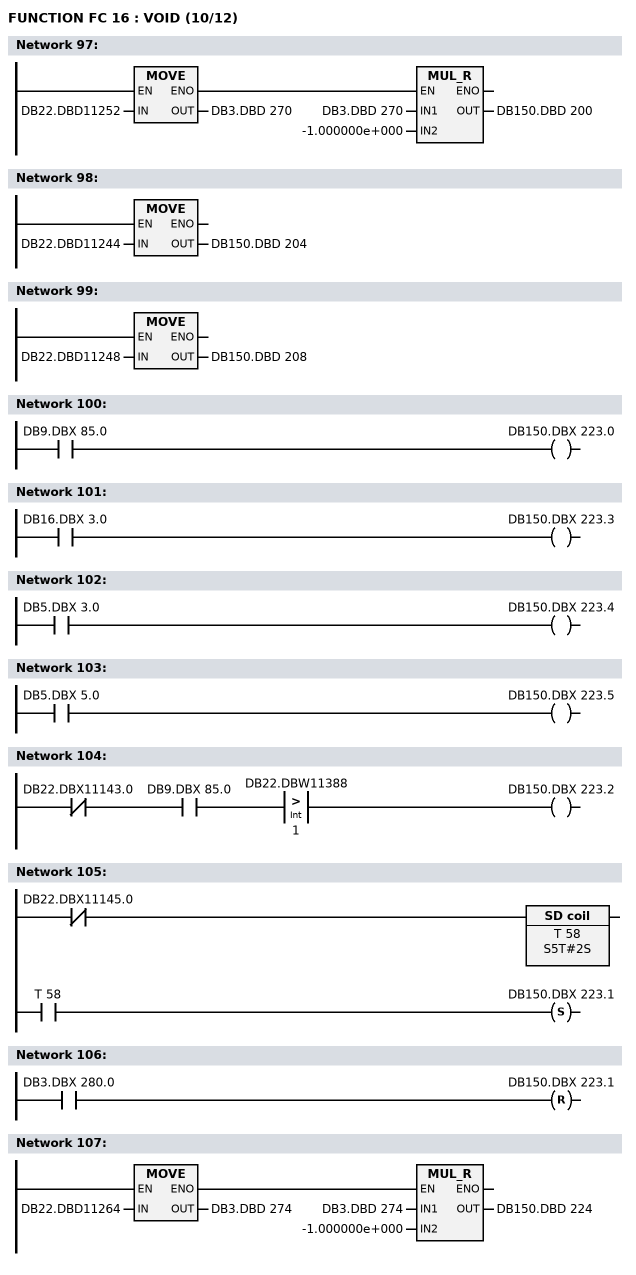

      A(    ;
      L     DB22.DBD11252;
      T     DB3.DBD  270;
      SET   ;
      SAVE  ;
      CLR   ;
      A     BR;
      )     ;
      JNB   M017;
      L     DB3.DBD  270;
      L     -1.000000e+000;
      *R    ;
      T     DB150.DBD  200;
M017: NOP   0;
NETWORK
TITLE =

      L     DB22.DBD11244;
      T     DB150.DBD  204;
      NOP   0;
NETWORK
TITLE =

      L     DB22.DBD11248;
      T     DB150.DBD  208;
      NOP   0;
NETWORK
TITLE =

      A     DB9.DBX   85.0;
      =     DB150.DBX  223.0;
NETWORK
TITLE =

      A     DB16.DBX    3.0;
      =     DB150.DBX  223.3;
NETWORK
TITLE =

      A     DB5.DBX    3.0;
      =     DB150.DBX  223.4;
NETWORK
TITLE =

      A     DB5.DBX    5.0;
      =     DB150.DBX  223.5;
NETWORK
TITLE =

      AN    DB22.DBX11143.0;
      A     DB9.DBX   85.0;
      A(    ;
      L     DB22.DBW11388;
      L     1;
      >I    ;
      )     ;
      =     DB150.DBX  223.2;
NETWORK
TITLE =

      AN    DB22.DBX11145.0;
      L     S5T#2S;
      SD    T     58;
      NOP   0;
      NOP   0;
      NOP   0;
      A     T     58;
      S     DB150.DBX  223.1;
NETWORK
TITLE =

      A     DB3.DBX  280.0;
      R     DB150.DBX  223.1;
NETWORK
TITLE =

      A(    ;
      L     DB22.DBD11264;
      T     DB3.DBD  274;
      SET   ;
      SAVE  ;
      CLR   ;
      A     BR;
      )     ;
      JNB   M018;
      L     DB3.DBD  274;
      L     -1.000000e+000;
      *R    ;
      T     DB150.DBD  224;
M018: NOP   0;
NETWORK
TITLE =
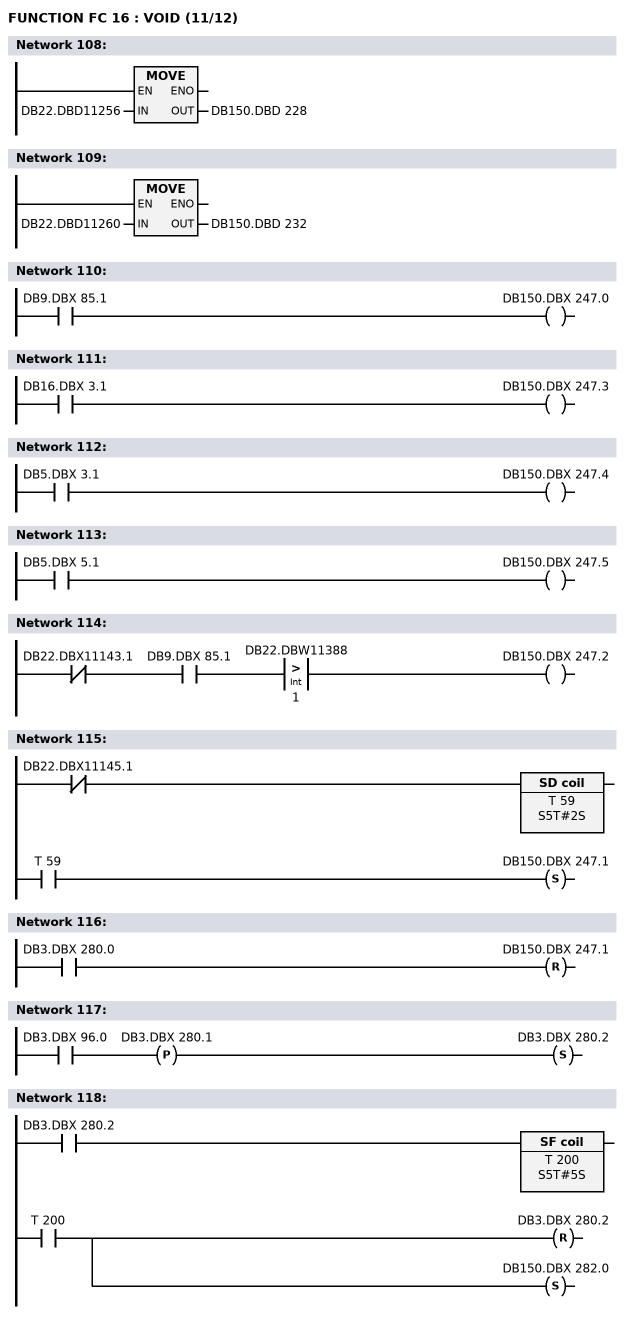

      L     DB22.DBD11256;
      T     DB150.DBD  228;
      NOP   0;
NETWORK
TITLE =

      L     DB22.DBD11260;
      T     DB150.DBD  232;
      NOP   0;
NETWORK
TITLE =

      A     DB9.DBX   85.1;
      =     DB150.DBX  247.0;
NETWORK
TITLE =

      A     DB16.DBX    3.1;
      =     DB150.DBX  247.3;
NETWORK
TITLE =

      A     DB5.DBX    3.1;
      =     DB150.DBX  247.4;
NETWORK
TITLE =

      A     DB5.DBX    5.1;
      =     DB150.DBX  247.5;
NETWORK
TITLE =

      AN    DB22.DBX11143.1;
      A     DB9.DBX   85.1;
      A(    ;
      L     DB22.DBW11388;
      L     1;
      >I    ;
      )     ;
      =     DB150.DBX  247.2;
NETWORK
TITLE =

      AN    DB22.DBX11145.1;
      L     S5T#2S;
      SD    T     59;
      NOP   0;
      NOP   0;
      NOP   0;
      A     T     59;
      S     DB150.DBX  247.1;
NETWORK
TITLE =

      A     DB3.DBX  280.0;
      R     DB150.DBX  247.1;
NETWORK
TITLE =

      A     DB3.DBX   96.0;
      BLD   100;
      FP    DB3.DBX  280.1;
      S     DB3.DBX  280.2;
NETWORK
TITLE =

      A     DB3.DBX  280.2;
      L     S5T#5S;
      SF    T    200;
      NOP   0;
      NOP   0;
      NOP   0;
      A     T    200;
      R     DB3.DBX  280.2;
      S     DB150.DBX  282.0;
NETWORK
TITLE =
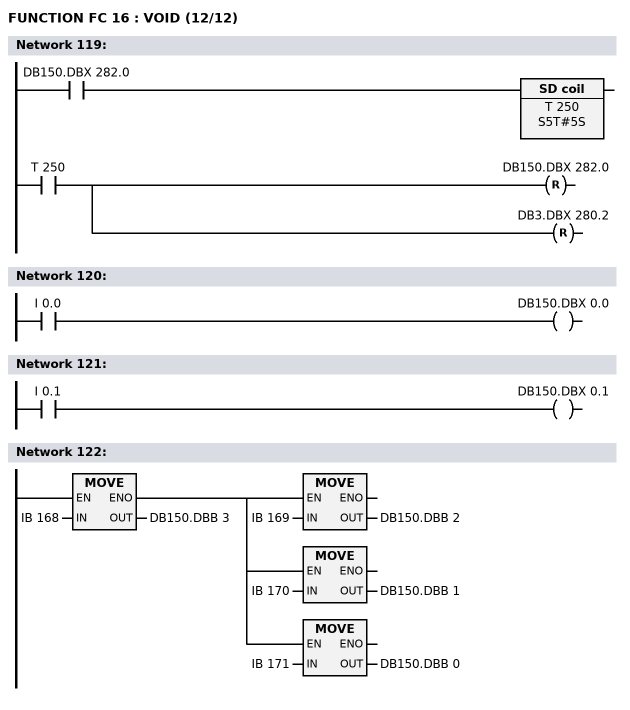

      A     DB150.DBX  282.0;
      L     S5T#5S;
      SD    T    250;
      NOP   0;
      NOP   0;
      NOP   0;
      A     T    250;
      R     DB150.DBX  282.0;
      R     DB3.DBX  280.2;
NETWORK
TITLE =

      A     I      0.0;
      =     DB150.DBX    0.0;
NETWORK
TITLE =

      A     I      0.1;
      =     DB150.DBX    0.1;
NETWORK
TITLE =

      L     IB   168;
      T     DB150.DBB    3;
      SET   ;
      SAVE  ;
      CLR   ;
      A     BR;
      =     L      0.0;
      A     L      0.0;
      JNB   M019;
      L     IB   169;
      T     DB150.DBB    2;
M019: NOP   0;
      A     L      0.0;
      JNB   M01a;
      L     IB   170;
      T     DB150.DBB    1;
M01a: NOP   0;
      A     L      0.0;
      JNB   M01b;
      L     IB   171;
      T     DB150.DBB    0;
M01b: NOP   0;
END_FUNCTION

DATA_BLOCK DB 250
VERSION : 0.0

 FB 250
BEGIN
   IN0 := 1;
   IN1 := W#16#180;
   IN2 := 95;
   IN3 := 95;
   OUT4 := FALSE;
   OUT5 := W#16#0;
   STAT6.STAT7 := W#16#64F1;
   STAT6.STAT8 := W#16#0;
   STAT6.STAT9 := W#16#61;
   STAT6.STAT10 := B#16#1;
   STAT6.STAT11 := B#16#3;
   STAT6.STAT12 := B#16#5E;
   STAT6.STAT13 := B#16#0;
   STAT6.STAT14 := B#16#2;
   STAT6.STAT15 := B#16#0;
   STAT6.STAT16 := B#16#0;
   STAT6.STAT17 := B#16#0;
   STAT6.STAT18 := B#16#0;
   STAT6.STAT19 := B#16#0;
   STAT6.STAT20 := B#16#0;
   STAT6.STAT21 := B#16#0;
   STAT6.STAT22 := B#16#0;
   STAT6.STAT23 := B#16#0;
   STAT6.STAT24 := B#16#0;
   STAT6.STAT25 := B#16#0;
   STAT6.STAT26 := B#16#0;
   STAT6.STAT27 := B#16#0;
   STAT6.STAT28 := B#16#0;
   STAT6.STAT29 := B#16#0;
   STAT6.STAT30 := B#16#0;
   STAT6.STAT31 := B#16#10;
   STAT6.STAT32 := B#16#C4;
   STAT6.STAT33 := B#16#D;
   STAT6.STAT34 := B#16#E6;
   STAT6.STAT35 := B#16#42;
   STAT6.STAT36 := B#16#43;
   STAT6.STAT37 := B#16#46;
   STAT6.STAT38 := B#16#49;
   STAT6.STAT39 := B#16#F5;
   STAT6.STAT40 := B#16#EC;
   STAT6.STAT41 := B#16#FA;
   STAT6.STAT42 := B#16#87;
   STAT6.STAT43 := B#16#F3;
   STAT6.STAT44 := B#16#C6;
   STAT6.STAT45 := B#16#F5;
   STAT6.STAT46 := B#16#F3;
   STAT6.STAT47 := B#16#0;
   STAT6.STAT48 := B#16#0;
   STAT6.STAT49 := B#16#0;
   STAT6.STAT50 := B#16#0;
   STAT6.STAT51 := B#16#F0;
   STAT6.STAT52 := B#16#99;
   STAT6.STAT53 := B#16#2E;
   STAT6.STAT54 := B#16#11;
   STAT6.STAT55 := B#16#EC;
   STAT6.STAT56 := B#16#26;
   STAT6.STAT57 := B#16#EA;
   STAT6.STAT58 := B#16#50;
   STAT6.STAT59 := B#16#ED;
   STAT6.STAT60 := B#16#65;
   STAT6.STAT61 := B#16#EB;
   STAT6.STAT62 := B#16#2;
   STAT6.STAT63 := B#16#5D;
   STAT6.STAT64 := B#16#22;
   STAT6.STAT65 := B#16#5E;
   STAT6.STAT66 := B#16#FF;
   STAT6.STAT67 := B#16#0;
   STAT6.STAT68 := B#16#0;
   STAT6.STAT69 := B#16#0;
   STAT6.STAT70 := B#16#0;
   STAT6.STAT71 := B#16#2;
   STAT6.STAT72 := B#16#0;
   STAT6.STAT73 := B#16#1C;
   STAT6.STAT74 := B#16#AA;
   STAT6.STAT75 := B#16#FE;
   STAT6.STAT76 := B#16#46;
   STAT6.STAT77 := B#16#FD;
   STAT6.STAT78 := B#16#61;
   STAT6.STAT79 := B#16#F8;
   STAT6.STAT80 := B#16#F9;
   STAT6.STAT81 := B#16#F8;
   STAT6.STAT82 := B#16#50;
   STAT6.STAT83 := B#16#49;
   STAT6.STAT84 := B#16#E1;
   STAT6.STAT85 := B#16#4B;
   STAT6.STAT86 := B#16#B0;
   STAT6.STAT87 := B#16#0;
   STAT6.STAT88 := B#16#0;
   STAT6.STAT89 := B#16#0;
   STAT6.STAT90 := B#16#0;
   STAT6.STAT91 := B#16#BB;
   STAT6.STAT92 := B#16#37;
   STAT6.STAT93 := B#16#63;
   STAT6.STAT94 := B#16#73;
   STAT6.STAT95 := B#16#A;
   STAT6.STAT96 := B#16#D1;
   STAT6.STAT97 := B#16#C;
   STAT6.STAT98 := B#16#2A;
   STAT6.STAT99 := B#16#E;
   STAT6.STAT100 := B#16#7E;
   STAT6.STAT101 := B#16#10;
   STAT6.STAT102 := B#16#2;
   STAT6.STAT103 := B#16#0;
   STAT6.STAT104 := B#16#19;
   STAT6.STAT105 := B#16#FD;
   STAT6.STAT106 := B#16#B6;
   STAT6.STAT107 := B#16#0;
   STAT6.STAT108 := B#16#0;
   STAT6.STAT109 := B#16#0;
   STAT6.STAT110 := B#16#0;
   STAT6.STAT111 := B#16#0;
   STAT6.STAT112 := B#16#0;
   STAT6.STAT113 := B#16#0;
   STAT6.STAT114 := B#16#0;
   STAT6.STAT115 := B#16#0;
   STAT6.STAT116 := B#16#0;
   STAT6.STAT117 := B#16#0;
   STAT6.STAT118 := B#16#0;
   STAT6.STAT119 := B#16#0;
   STAT6.STAT120 := B#16#0;
   STAT6.STAT121 := B#16#0;
   STAT6.STAT122 := B#16#0;
   STAT6.STAT123 := B#16#0;
   STAT6.STAT124 := B#16#0;
   STAT6.STAT125 := B#16#0;
   STAT6.STAT126 := B#16#0;
   STAT6.STAT127 := B#16#0;
   STAT6.STAT128 := B#16#0;
   STAT6.STAT129 := B#16#0;
   STAT6.STAT130 := B#16#0;
   STAT6.STAT131 := B#16#0;
   STAT6.STAT132 := B#16#0;
   STAT6.STAT133 := B#16#0;
   STAT6.STAT134 := B#16#0;
   STAT6.STAT135 := B#16#0;
   STAT6.STAT136 := B#16#0;
   STAT6.STAT137 := B#16#0;
   STAT6.STAT138 := B#16#0;
   STAT6.STAT139 := B#16#0;
   STAT6.STAT140 := B#16#0;
   STAT6.STAT141 := B#16#0;
   STAT6.STAT142 := B#16#0;
   STAT6.STAT143 := B#16#0;
   STAT6.STAT144 := B#16#0;
   STAT6.STAT145 := B#16#0;
   STAT6.STAT146 := B#16#0;
   STAT6.STAT147 := B#16#0;
   STAT6.STAT148 := B#16#0;
   STAT6.STAT149 := B#16#0;
   STAT6.STAT150 := B#16#0;
   STAT6.STAT151 := B#16#0;
   STAT6.STAT152 := B#16#0;
   STAT6.STAT153 := B#16#0;
   STAT6.STAT154 := B#16#0;
   STAT6.STAT155 := B#16#0;
   STAT6.STAT156 := B#16#0;
   STAT6.STAT157 := B#16#0;
   STAT6.STAT158 := B#16#0;
   STAT6.STAT159 := B#16#0;
   STAT6.STAT160 := B#16#0;
   STAT6.STAT161 := B#16#0;
   STAT6.STAT162 := B#16#0;
   STAT6.STAT163 := B#16#0;
   STAT6.STAT164 := B#16#0;
   STAT6.STAT165 := B#16#0;
   STAT6.STAT166 := B#16#0;
   STAT6.STAT167 := B#16#0;
   STAT6.STAT168 := B#16#0;
   STAT6.STAT169 := B#16#0;
   STAT6.STAT170 := B#16#0;
   STAT6.STAT171 := B#16#0;
   STAT6.STAT172 := B#16#0;
   STAT6.STAT173 := B#16#0;
   STAT6.STAT174 := B#16#0;
   STAT6.STAT175 := B#16#0;
   STAT6.STAT176 := B#16#0;
   STAT6.STAT177 := B#16#0;
   STAT6.STAT178 := B#16#0;
   STAT6.STAT179 := B#16#0;
   STAT6.STAT180 := B#16#0;
   STAT6.STAT181 := B#16#0;
   STAT6.STAT182 := B#16#0;
   STAT6.STAT183 := B#16#0;
   STAT6.STAT184 := B#16#0;
   STAT6.STAT185 := B#16#0;
   STAT6.STAT186 := B#16#0;
   STAT6.STAT187 := B#16#0;
   STAT6.STAT188 := B#16#0;
   STAT6.STAT189 := B#16#0;
   STAT6.STAT190 := B#16#0;
   STAT6.STAT191 := B#16#0;
   STAT6.STAT192 := B#16#0;
   STAT6.STAT193 := B#16#0;
   STAT6.STAT194 := B#16#0;
   STAT6.STAT195 := B#16#0;
   STAT6.STAT196 := B#16#0;
   STAT6.STAT197 := B#16#0;
   STAT6.STAT198 := B#16#0;
   STAT6.STAT199 := B#16#0;
   STAT6.STAT200 := B#16#0;
   STAT6.STAT201 := B#16#0;
   STAT6.STAT202 := B#16#0;
   STAT6.STAT203 := B#16#0;
   STAT6.STAT204 := B#16#0;
   STAT6.STAT205 := B#16#0;
   STAT6.STAT206 := B#16#0;
   STAT6.STAT207 := B#16#0;
   STAT6.STAT208 := B#16#0;
   STAT6.STAT209 := B#16#0;
   STAT6.STAT210 := B#16#0;
   STAT6.STAT211 := B#16#0;
   STAT6.STAT212 := B#16#0;
   STAT6.STAT213 := B#16#0;
   STAT6.STAT214 := B#16#0;
   STAT6.STAT215 := B#16#0;
   STAT6.STAT216 := B#16#0;
   STAT6.STAT217 := B#16#0;
   STAT6.STAT218 := B#16#0;
   STAT6.STAT219 := B#16#0;
   STAT6.STAT220 := B#16#0;
   STAT6.STAT221 := B#16#0;
   STAT6.STAT222 := B#16#0;
   STAT6.STAT223 := B#16#0;
   STAT6.STAT224 := B#16#0;
   STAT6.STAT225 := B#16#0;
   STAT6.STAT226 := B#16#0;
   STAT6.STAT227 := B#16#0;
   STAT6.STAT228 := B#16#0;
   STAT6.STAT229 := B#16#0;
   STAT6.STAT230 := B#16#0;
   STAT6.STAT231 := B#16#0;
   STAT6.STAT232 := B#16#0;
   STAT6.STAT233 := B#16#0;
   STAT6.STAT234 := B#16#0;
   STAT6.STAT235 := B#16#0;
   STAT6.STAT236 := B#16#0;
   STAT6.STAT237 := B#16#0;
   STAT6.STAT238 := B#16#0;
   STAT6.STAT239 := B#16#0;
   STAT6.STAT240 := B#16#0;
   STAT6.STAT241 := B#16#0;
   STAT6.STAT242 := B#16#0;
   STAT6.STAT243 := B#16#0;
   STAT6.STAT244 := B#16#0;
   STAT6.STAT245 := B#16#0;
   STAT6.STAT246 := B#16#0;
   STAT6.STAT247 := B#16#0;
   STAT6.STAT248 := B#16#0;
   STAT6.STAT249 := B#16#0;
   STAT6.STAT250 := B#16#0;
   STAT6.STAT251 := B#16#0;
   STAT6.STAT252 := B#16#0;
   STAT6.STAT253 := B#16#0;
   STAT6.STAT254 := B#16#0;
   STAT6.STAT255 := B#16#0;
   STAT6.STAT256 := B#16#0;
   STAT6.STAT257 := B#16#0;
   STAT6.STAT258 := B#16#0;
   STAT6.STAT259 := B#16#0;
   STAT6.STAT260 := B#16#0;
   STAT261.STAT262 := W#16#64F1;
   STAT261.STAT263 := W#16#0;
   STAT261.STAT264 := W#16#6;
   STAT261.STAT265 := B#16#1;
   STAT261.STAT266 := B#16#3;
   STAT261.STAT267 := W#16#0;
   STAT261.STAT268 := W#16#2F;
   STAT261.STAT269 := B#16#0;
   STAT261.STAT270 := B#16#0;
   STAT261.STAT271 := B#16#0;
   STAT261.STAT272 := B#16#0;
   STAT261.STAT273 := B#16#0;
   STAT261.STAT274 := B#16#0;
   STAT261.STAT275 := B#16#0;
   STAT261.STAT276 := B#16#0;
   STAT261.STAT277 := B#16#0;
   STAT261.STAT278 := B#16#0;
   STAT261.STAT279 := B#16#0;
   STAT261.STAT280 := B#16#0;
   STAT261.STAT281 := B#16#0;
   STAT261.STAT282 := B#16#0;
   STAT261.STAT283 := B#16#0;
   STAT261.STAT284 := B#16#0;
   STAT261.STAT285 := B#16#0;
   STAT261.STAT286 := B#16#0;
   STAT261.STAT287 := B#16#0;
   STAT261.STAT288 := B#16#0;
   STAT261.STAT289 := B#16#0;
   STAT261.STAT290 := B#16#0;
   STAT261.STAT291 := B#16#0;
   STAT261.STAT292 := B#16#0;
   STAT261.STAT293 := B#16#0;
   STAT261.STAT294 := B#16#0;
   STAT261.STAT295 := B#16#0;
   STAT261.STAT296 := B#16#0;
   STAT261.STAT297 := B#16#0;
   STAT261.STAT298 := B#16#0;
   STAT261.STAT299 := B#16#0;
   STAT261.STAT300 := B#16#0;
   STAT261.STAT301 := B#16#0;
   STAT261.STAT302 := B#16#0;
   STAT261.STAT303 := B#16#0;
   STAT261.STAT304 := B#16#0;
   STAT261.STAT305 := B#16#0;
   STAT261.STAT306 := B#16#0;
   STAT261.STAT307 := B#16#0;
   STAT261.STAT308 := B#16#0;
   STAT261.STAT309 := B#16#0;
   STAT261.STAT310 := B#16#0;
   STAT261.STAT311 := B#16#0;
   STAT261.STAT312 := B#16#0;
   STAT261.STAT313 := B#16#0;
   STAT261.STAT314 := B#16#0;
   STAT261.STAT315 := B#16#0;
   STAT261.STAT316 := B#16#0;
   STAT261.STAT317 := B#16#0;
   STAT261.STAT318 := B#16#0;
   STAT261.STAT319 := B#16#0;
   STAT261.STAT320 := B#16#0;
   STAT261.STAT321 := B#16#0;
   STAT261.STAT322 := B#16#0;
   STAT261.STAT323 := B#16#0;
   STAT261.STAT324 := B#16#0;
   STAT261.STAT325 := B#16#0;
   STAT261.STAT326 := B#16#0;
   STAT261.STAT327 := B#16#0;
   STAT261.STAT328 := B#16#0;
   STAT261.STAT329 := B#16#0;
   STAT261.STAT330 := B#16#0;
   STAT261.STAT331 := B#16#0;
   STAT261.STAT332 := B#16#0;
   STAT261.STAT333 := B#16#0;
   STAT261.STAT334 := B#16#0;
   STAT261.STAT335 := B#16#0;
   STAT261.STAT336 := B#16#0;
   STAT261.STAT337 := B#16#0;
   STAT261.STAT338 := B#16#0;
   STAT261.STAT339 := B#16#0;
   STAT261.STAT340 := B#16#0;
   STAT261.STAT341 := B#16#0;
   STAT261.STAT342 := B#16#0;
   STAT261.STAT343 := B#16#0;
   STAT261.STAT344 := B#16#0;
   STAT261.STAT345 := B#16#0;
   STAT261.STAT346 := B#16#0;
   STAT261.STAT347 := B#16#0;
   STAT261.STAT348 := B#16#0;
   STAT261.STAT349 := B#16#0;
   STAT261.STAT350 := B#16#0;
   STAT261.STAT351 := B#16#0;
   STAT261.STAT352 := B#16#0;
   STAT261.STAT353 := B#16#0;
   STAT261.STAT354 := B#16#0;
   STAT261.STAT355 := B#16#0;
   STAT261.STAT356 := B#16#0;
   STAT261.STAT357 := B#16#0;
   STAT261.STAT358 := B#16#0;
   STAT261.STAT359 := B#16#0;
   STAT261.STAT360 := B#16#0;
   STAT261.STAT361 := B#16#0;
   STAT261.STAT362 := B#16#0;
   STAT261.STAT363 := B#16#0;
   STAT261.STAT364 := B#16#0;
   STAT261.STAT365 := B#16#0;
   STAT261.STAT366 := B#16#0;
   STAT261.STAT367 := B#16#0;
   STAT261.STAT368 := B#16#0;
   STAT261.STAT369 := B#16#0;
   STAT261.STAT370 := B#16#0;
   STAT261.STAT371 := B#16#0;
   STAT261.STAT372 := B#16#0;
   STAT261.STAT373 := B#16#0;
   STAT261.STAT374 := B#16#0;
   STAT261.STAT375 := B#16#0;
   STAT261.STAT376 := B#16#0;
   STAT261.STAT377 := B#16#0;
   STAT261.STAT378 := B#16#0;
   STAT261.STAT379 := B#16#0;
   STAT261.STAT380 := B#16#0;
   STAT261.STAT381 := B#16#0;
   STAT261.STAT382 := B#16#0;
   STAT261.STAT383 := B#16#0;
   STAT261.STAT384 := B#16#0;
   STAT261.STAT385 := B#16#0;
   STAT261.STAT386 := B#16#0;
   STAT261.STAT387 := B#16#0;
   STAT261.STAT388 := B#16#0;
   STAT261.STAT389 := B#16#0;
   STAT261.STAT390 := B#16#0;
   STAT261.STAT391 := B#16#0;
   STAT261.STAT392 := B#16#0;
   STAT261.STAT393 := B#16#0;
   STAT261.STAT394 := B#16#0;
   STAT261.STAT395 := B#16#0;
   STAT261.STAT396 := B#16#0;
   STAT261.STAT397 := B#16#0;
   STAT261.STAT398 := B#16#0;
   STAT261.STAT399 := B#16#0;
   STAT261.STAT400 := B#16#0;
   STAT261.STAT401 := B#16#0;
   STAT261.STAT402 := B#16#0;
   STAT261.STAT403 := B#16#0;
   STAT261.STAT404 := B#16#0;
   STAT261.STAT405 := B#16#0;
   STAT261.STAT406 := B#16#0;
   STAT261.STAT407 := B#16#0;
   STAT261.STAT408 := B#16#0;
   STAT261.STAT409 := B#16#0;
   STAT261.STAT410 := B#16#0;
   STAT261.STAT411 := B#16#0;
   STAT261.STAT412 := B#16#0;
   STAT261.STAT413 := B#16#0;
   STAT261.STAT414 := B#16#0;
   STAT261.STAT415 := B#16#0;
   STAT261.STAT416 := B#16#0;
   STAT261.STAT417 := B#16#0;
   STAT261.STAT418 := B#16#0;
   STAT261.STAT419 := B#16#0;
   STAT261.STAT420 := B#16#0;
   STAT261.STAT421 := B#16#0;
   STAT261.STAT422 := B#16#0;
   STAT261.STAT423 := B#16#0;
   STAT261.STAT424 := B#16#0;
   STAT261.STAT425 := B#16#0;
   STAT261.STAT426 := B#16#0;
   STAT261.STAT427 := B#16#0;
   STAT261.STAT428 := B#16#0;
   STAT261.STAT429 := B#16#0;
   STAT261.STAT430 := B#16#0;
   STAT261.STAT431 := B#16#0;
   STAT261.STAT432 := B#16#0;
   STAT261.STAT433 := B#16#0;
   STAT261.STAT434 := B#16#0;
   STAT261.STAT435 := B#16#0;
   STAT261.STAT436 := B#16#0;
   STAT261.STAT437 := B#16#0;
   STAT261.STAT438 := B#16#0;
   STAT261.STAT439 := B#16#0;
   STAT261.STAT440 := B#16#0;
   STAT261.STAT441 := B#16#0;
   STAT261.STAT442 := B#16#0;
   STAT261.STAT443 := B#16#0;
   STAT261.STAT444 := B#16#0;
   STAT261.STAT445 := B#16#0;
   STAT261.STAT446 := B#16#0;
   STAT261.STAT447 := B#16#0;
   STAT261.STAT448 := B#16#0;
   STAT261.STAT449 := B#16#0;
   STAT261.STAT450 := B#16#0;
   STAT261.STAT451 := B#16#0;
   STAT261.STAT452 := B#16#0;
   STAT261.STAT453 := B#16#0;
   STAT261.STAT454 := B#16#0;
   STAT261.STAT455 := B#16#0;
   STAT261.STAT456 := B#16#0;
   STAT261.STAT457 := B#16#0;
   STAT261.STAT458 := B#16#0;
   STAT261.STAT459 := B#16#0;
   STAT261.STAT460 := B#16#0;
   STAT261.STAT461 := B#16#0;
   STAT261.STAT462 := B#16#0;
   STAT261.STAT463 := B#16#0;
   STAT261.STAT464 := B#16#0;
   STAT261.STAT465 := B#16#0;
   STAT261.STAT466 := B#16#0;
   STAT261.STAT467 := B#16#0;
   STAT261.STAT468 := B#16#0;
   STAT261.STAT469 := B#16#0;
   STAT261.STAT470 := B#16#0;
   STAT261.STAT471 := B#16#0;
   STAT261.STAT472 := B#16#0;
   STAT261.STAT473 := B#16#0;
   STAT261.STAT474 := B#16#0;
   STAT261.STAT475 := B#16#0;
   STAT261.STAT476 := B#16#0;
   STAT261.STAT477 := B#16#0;
   STAT261.STAT478 := B#16#0;
   STAT261.STAT479 := B#16#0;
   STAT261.STAT480 := B#16#0;
   STAT261.STAT481 := B#16#0;
   STAT261.STAT482 := B#16#0;
   STAT261.STAT483 := B#16#0;
   STAT261.STAT484 := B#16#0;
   STAT261.STAT485 := B#16#0;
   STAT261.STAT486 := B#16#0;
   STAT261.STAT487 := B#16#0;
   STAT261.STAT488 := B#16#0;
   STAT261.STAT489 := B#16#0;
   STAT261.STAT490 := B#16#0;
   STAT261.STAT491 := B#16#0;
   STAT261.STAT492 := B#16#0;
   STAT261.STAT493 := B#16#0;
   STAT261.STAT494 := B#16#0;
   STAT261.STAT495 := B#16#0;
   STAT261.STAT496 := B#16#0;
   STAT261.STAT497 := B#16#0;
   STAT261.STAT498 := B#16#0;
   STAT261.STAT499 := B#16#0;
   STAT261.STAT500 := B#16#0;
   STAT261.STAT501 := B#16#0;
   STAT261.STAT502 := B#16#0;
   STAT261.STAT503 := B#16#0;
   STAT261.STAT504 := B#16#0;
   STAT261.STAT505 := B#16#0;
   STAT261.STAT506 := B#16#0;
   STAT261.STAT507 := B#16#0;
   STAT261.STAT508 := B#16#0;
   STAT261.STAT509 := B#16#0;
   STAT261.STAT510 := B#16#0;
   STAT261.STAT511 := B#16#0;
   STAT261.STAT512 := B#16#0;
   STAT261.STAT513 := B#16#0;
   STAT261.STAT514 := B#16#0;
   STAT515 := 0;
   STAT516 := 0;
   STAT517 := TRUE;
   STAT518 := FALSE;
   STAT519 := FALSE;
   STAT520 := FALSE;
   STAT521 := W#16#8180;
   STAT522 := 0;
   STAT523 := TRUE;
   STAT524 := FALSE;
   STAT525 := W#16#0;
   STAT526 := 6;
   STAT527 := 103;
   STAT528 := FALSE;
   STAT529 := FALSE;
   STAT530 := W#16#0;
   STAT531 := FALSE;
   STAT532 := W#16#1;
   STAT533.IN := FALSE;
   STAT533.PT := T#0MS;
   STAT533.Q := FALSE;
   STAT533.ET := T#0MS;
   STAT533.STATE := B#16#0;
   STAT533.STIME := T#0MS;
   STAT533.ATIME := T#0MS;
   STAT541 := FALSE;
   STAT542 := FALSE;
   STAT543 := FALSE;
   STAT544 := W#16#0;
END_DATA_BLOCK

ORGANIZATION_BLOCK OB 82
VERSION : 0.1


VAR_TEMP
  TEMP0 : BYTE ;
  TEMP1 : BYTE ;
  TEMP2 : BYTE ;
  TEMP3 : BYTE ;
  TEMP4 : BYTE ;
  TEMP5 : BYTE ;
  TEMP6 : WORD ;
  TEMP7 : BOOL ;
  TEMP8 : BOOL ;
  TEMP9 : BOOL ;
  TEMP10 : BOOL ;
  TEMP11 : BOOL ;
  TEMP12 : BOOL ;
  TEMP13 : BOOL ;
  TEMP14 : BOOL ;
  TEMP15 : BYTE ;
  TEMP16 : BOOL ;
  TEMP17 : BOOL ;
  TEMP18 : BOOL ;
  TEMP19 : BOOL ;
  TEMP20 : BOOL ;
  TEMP21 : BOOL ;
  TEMP22 : BOOL ;
  TEMP23 : BOOL ;
  TEMP24 : BOOL ;
  TEMP25 : BOOL ;
  TEMP26 : BOOL ;
  TEMP27 : BOOL ;
  TEMP28 : BOOL ;
  TEMP29 : BOOL ;
  TEMP30 : BOOL ;
  TEMP31 : BOOL ;
  TEMP32 : DATE_AND_TIME ;
END_VAR
BEGIN
NETWORK
TITLE =

END_ORGANIZATION_BLOCK

ORGANIZATION_BLOCK OB 85
VERSION : 0.1


VAR_TEMP
  TEMP0 : BYTE ;
  TEMP1 : BYTE ;
  TEMP2 : BYTE ;
  TEMP3 : BYTE ;
  TEMP4 : BYTE ;
  TEMP5 : BYTE ;
  TEMP6 : INT ;
  TEMP7 : BYTE ;
  TEMP8 : BYTE ;
  TEMP9 : BYTE ;
  TEMP10 : BYTE ;
  TEMP11 : DATE_AND_TIME ;
END_VAR
BEGIN
NETWORK
TITLE =

END_ORGANIZATION_BLOCK

ORGANIZATION_BLOCK OB 86
VERSION : 0.1


VAR_TEMP
  TEMP0 : BYTE ;
  TEMP1 : BYTE ;
  TEMP2 : BYTE ;
  TEMP3 : BYTE ;
  TEMP4 : BYTE ;
  TEMP5 : BYTE ;
  TEMP6 : WORD ;
  TEMP7 : ARRAY  [0 .. 31 ] OF BOOL ;
  TEMP8 : DATE_AND_TIME ;
END_VAR
BEGIN
NETWORK
TITLE =

END_ORGANIZATION_BLOCK

ORGANIZATION_BLOCK OB 122
VERSION : 0.1


VAR_TEMP
  TEMP0 : BYTE ;
  TEMP1 : BYTE ;
  TEMP2 : BYTE ;
  TEMP3 : BYTE ;
  TEMP4 : BYTE ;
  TEMP5 : BYTE ;
  TEMP6 : WORD ;
  TEMP7 : WORD ;
  TEMP8 : WORD ;
  TEMP9 : DATE_AND_TIME ;
END_VAR
BEGIN
NETWORK
TITLE =

END_ORGANIZATION_BLOCK

